FUNCTION_BLOCK FB_MqttLightProtocol
VAR_INPUT
    bTestNamespace : BOOL := FALSE;
    bCatalogReady : BOOL := TRUE;
    nLightCount : DINT := -1;
END_VAR
VAR_OUTPUT
    nCount : UINT;
    nRejectedQueue : UDINT;
    nRejectedInput : UDINT;
    bReady : BOOL;
    nStateIndex : DINT;
    sStateTopic : STRING(255);
    sStatePayload : STRING(3);
    bPublishPending : BOOL;
END_VAR
VAR
    aQueue : ARRAY[1..16] OF ST_LightCommand;
    nHead : UINT := 1;
    aSentTopic : ARRAY[1..16] OF STRING(255);
    aSentOn : ARRAY[1..16] OF BOOL;
    aSentValid : ARRAY[1..16] OF BOOL;
    nPendingIndex : DINT;
    sPendingTopic : STRING(255);
    bPendingOn : BOOL;
    fbTopicMap : FB_MqttTopicMap;
END_VAR

METHOD PUBLIC Reset
VAR
    i : UINT;
END_VAR
nHead := 1;
nCount := 0;
bPublishPending := FALSE;
nPendingIndex := 0;
FOR i := 1 TO 16 DO
    aQueue[i].bValid := FALSE;
    aSentValid[i] := FALSE;
END_FOR
END_METHOD

METHOD PUBLIC RequestSnapshot
VAR
    i : UINT;
END_VAR
FOR i := 1 TO 16 DO
    aSentValid[i] := FALSE;
END_FOR
bPublishPending := FALSE;
nPendingIndex := 0;
END_METHOD

METHOD PUBLIC SetConnection
VAR_INPUT
    bNewReady : BOOL;
END_VAR
VAR
    i : UINT;
END_VAR
IF (bNewReady <> bReady) OR NOT bNewReady THEN
    nHead := 1;
    nCount := 0;
    FOR i := 1 TO 16 DO
        aQueue[i].bValid := FALSE;
    END_FOR
END_IF
bReady := bNewReady;
END_METHOD

METHOD PUBLIC BuildTopic : STRING(255)
VAR_INPUT
    sLocationId : STRING(16);
    sLightId : STRING(16);
    sSuffix : STRING(8);
END_VAR
BuildTopic := fbTopicMap.BuildLightTopic(bTestNamespace := bTestNamespace, sLocationId := sLocationId, sLightId := sLightId, sSuffix := sSuffix);
END_METHOD

METHOD PUBLIC Receive : BOOL
VAR_INPUT
    sTopic : STRING(255);
    sPayload : STRING(8);
    nPayloadSize : UDINT;
END_VAR
VAR_IN_OUT
    aLights : ARRAY[*] OF ST_LightInfo;
END_VAR
VAR
    i : DINT;
    nActiveCount : DINT;
    nTail : UINT;

    bTargetOn : BOOL;
END_VAR
Receive := FALSE;
IF NOT bCatalogReady THEN
    nRejectedInput := nRejectedInput + 1;
    RETURN;
END_IF
nActiveCount := nLightCount;
IF nActiveCount = -1 THEN
    nActiveCount := UPPER_BOUND(aLights, 1) - LOWER_BOUND(aLights, 1) + 1;
END_IF
IF (nActiveCount < 0) OR (nActiveCount > 16) OR (nActiveCount > UPPER_BOUND(aLights, 1) - LOWER_BOUND(aLights, 1) + 1) THEN
    nRejectedInput := nRejectedInput + 1;
    RETURN;
END_IF
IF NOT bReady OR (nPayloadSize <> INT_TO_UDINT(LEN(sPayload))) THEN
    nRejectedInput := nRejectedInput + 1;
    RETURN;
END_IF
IF (sPayload = 'ON') AND (nPayloadSize = 2) THEN
    bTargetOn := TRUE;
ELSIF (sPayload = 'OFF') AND (nPayloadSize = 3) THEN
    bTargetOn := FALSE;
ELSE
    nRejectedInput := nRejectedInput + 1;
    RETURN;
END_IF
IF nActiveCount = 0 THEN
    nRejectedInput := nRejectedInput + 1;
    RETURN;
END_IF
FOR i := LOWER_BOUND(aLights, 1) TO LOWER_BOUND(aLights, 1) + nActiveCount - 1 DO
    IF sTopic = BuildTopic(sLocationId := aLights[i].sLocationId, sLightId := aLights[i].sId, sSuffix := 'set') THEN
        IF nCount >= 16 THEN
            nRejectedQueue := nRejectedQueue + 1;
            RETURN;
        END_IF
        nTail := nHead + nCount;
        IF nTail > 16 THEN
            nTail := nTail - 16;
        END_IF
        aQueue[nTail].sLocationId := aLights[i].sLocationId;
        aQueue[nTail].sLightId := aLights[i].sId;
        aQueue[nTail].bTargetOn := bTargetOn;
        aQueue[nTail].bValid := TRUE;
        nCount := nCount + 1;
        Receive := TRUE;
        RETURN;
    END_IF
END_FOR
nRejectedInput := nRejectedInput + 1;
END_METHOD

METHOD PUBLIC Pop : ST_LightCommand
Pop.bValid := FALSE;
IF bReady AND (nCount > 0) THEN
    Pop := aQueue[nHead];
    aQueue[nHead].bValid := FALSE;
    nHead := nHead + 1;
    IF nHead > 16 THEN
        nHead := 1;
    END_IF
    nCount := nCount - 1;
END_IF
END_METHOD

METHOD PUBLIC PlanState
VAR_IN_OUT
    aLights : ARRAY[*] OF ST_LightInfo;
END_VAR
VAR
    i : DINT;
    nSlot : DINT;
    nActiveCount : DINT;
END_VAR
bPublishPending := FALSE;
nStateIndex := 0;
sStateTopic := '';
sStatePayload := '';
IF NOT bCatalogReady THEN
    RETURN;
END_IF
nActiveCount := nLightCount;
IF nActiveCount = -1 THEN
    nActiveCount := UPPER_BOUND(aLights, 1) - LOWER_BOUND(aLights, 1) + 1;
END_IF
IF (nActiveCount < 0) OR (nActiveCount > 16) OR (nActiveCount > UPPER_BOUND(aLights, 1) - LOWER_BOUND(aLights, 1) + 1) OR (nActiveCount = 0) THEN
    RETURN;
END_IF
FOR i := LOWER_BOUND(aLights, 1) TO LOWER_BOUND(aLights, 1) + nActiveCount - 1 DO
    nSlot := i - LOWER_BOUND(aLights, 1) + 1;
    IF NOT aSentValid[nSlot] OR (aSentTopic[nSlot] <> BuildTopic(sLocationId := aLights[i].sLocationId, sLightId := aLights[i].sId, sSuffix := 'state')) OR (aSentOn[nSlot] <> aLights[i].bOn) THEN
        nStateIndex := i;
        sStateTopic := BuildTopic(sLocationId := aLights[i].sLocationId, sLightId := aLights[i].sId, sSuffix := 'state');
        IF aLights[i].bOn THEN
            sStatePayload := 'ON';
        ELSE
            sStatePayload := 'OFF';
        END_IF
        nPendingIndex := nSlot;
        sPendingTopic := sStateTopic;
        bPendingOn := aLights[i].bOn;
        bPublishPending := TRUE;
        RETURN;
    END_IF
END_FOR
END_METHOD

METHOD PUBLIC ConfirmPublish
VAR_INPUT
    bAccepted : BOOL;
END_VAR
IF bPublishPending AND bAccepted THEN
    aSentTopic[nPendingIndex] := sPendingTopic;
    aSentOn[nPendingIndex] := bPendingOn;
    aSentValid[nPendingIndex] := TRUE;
END_IF
bPublishPending := FALSE;
nPendingIndex := 0;
END_METHOD

END_FUNCTION_BLOCK

(* stored: Version 1.1.0.1
   POU FB_MqttLightProtocol: Id {b18f36f3-fcf2-4122-8e1a-67e1d0d90b21}, SpecialFunc None
   Method Reset: Id {c6b8309b-460b-4f70-b769-36e11ca7be5c}
   Method RequestSnapshot: Id {e128e520-4cb2-4c8f-91ee-f53ab81f013d}
   Method SetConnection: Id {fa095f20-95fd-43e8-8b11-4914a0d583e9}
   Method BuildTopic: Id {eef997cf-d1dd-4653-9437-99d271bfc2b5}
   Method Receive: Id {7d87b4c7-12e3-47a8-83c4-9e958d73c555}
   Method Pop: Id {be83d102-31ee-4367-9d51-aa8508a5ce89}
   Method PlanState: Id {169aeef9-0491-4bd2-8da2-c12b9a996ba8}
   Method ConfirmPublish: Id {0eeb70fd-150b-424f-a316-e5e20c347fd2} *)
